(* IEC 61131-3 sources: moqui-plc/rust-plc/interfaces/plcopen-motion, 3 files *)

(* ---- types.st ---- *)
(* PLCopen Motion Control - data types used by moqui-plc.
 *
 * Interface declarations only, for type checking with a non-CODESYS compiler.
 * Names follow PLCopen Motion Control Part 1 (single axis) and Part 4
 * (coordinated motion), with the enumeration spellings used in the canonical
 * iec61131 tree. A runtime that hosts moqui-plc provides the real types.
 *
 * AXIS_REF and AXES_GROUP_REF are opaque in PLCopen; the members below are the
 * only ones the moqui-plc code reads.
 *)

TYPE AXIS_REF :
STRUCT
    wDriveId : WORD; (* drive identifier, used for log naming *)
    fTaskCycle : LREAL; (* cycle time of the motion task that runs the axis [s] *)
END_STRUCT
END_TYPE

TYPE AXES_GROUP_REF :
STRUCT
    nAxes : INT;
END_STRUCT
END_TYPE

TYPE TRIGGER_REF :
STRUCT
    iTriggerNumber : INT;
END_STRUCT
END_TYPE

TYPE MC_BUFFER_MODE : (aborting, Buffered, BlendingLow, BlendingPrevious, BlendingNext, BlendingHigh); END_TYPE
TYPE MC_DIRECTION : (negative := -1, shortest, positive, current, fastest); END_TYPE
TYPE MC_STARTMODE : (absolute, relative, ramp_in); END_TYPE
TYPE MC_TRANSITION_MODE : (TMNone, TMStartVelocity, TMConstantVelocity, TMCornerDistance, TMMaxCornerDeviation); END_TYPE
TYPE MC_CIRC_PATHCHOICE : (CLOCKWISE, COUNTER_CLOCKWISE); END_TYPE

TYPE MC_COORD_REF :
STRUCT
    X : LREAL;
    Y : LREAL;
    Z : LREAL;
    A : LREAL;
    B : LREAL;
    C : LREAL;
END_STRUCT
END_TYPE

(* Profile and cam references: content is runtime specific. *)
TYPE MC_TP_REF : STRUCT nPoints : INT; END_STRUCT END_TYPE
TYPE MC_TV_REF : STRUCT nPoints : INT; END_STRUCT END_TYPE
TYPE MC_TA_REF : STRUCT nPoints : INT; END_STRUCT END_TYPE
TYPE MC_CAM_REF : STRUCT nElements : INT; END_STRUCT END_TYPE
TYPE MC_CAM_ID : STRUCT nId : UDINT; END_STRUCT END_TYPE

(* ---- part1-single-axis.st ---- *)
(* PLCopen Motion Control Part 1 - single-axis function blocks used by moqui-plc.
 *
 * Interface declarations only (no implementation), for type checking with a
 * non-CODESYS compiler. Parameters follow the PLCopen function block
 * interface; MC_Power also carries the drive-start and regulator inputs
 * the moqui-plc code sets.
 * A runtime that hosts moqui-plc implements these blocks with the same
 * signatures.
 *)

FUNCTION_BLOCK MC_Power
VAR_IN_OUT
    Axis : AXIS_REF;
END_VAR
VAR_INPUT
    Enable : BOOL;
    bRegulatorOn : BOOL;
    bDriveStart : BOOL;
END_VAR
VAR_OUTPUT
    Status : BOOL;
    bRegulatorRealState : BOOL;
    bDriveStartRealState : BOOL;
    Busy : BOOL;
    Error : BOOL;
    ErrorID : WORD;
END_VAR
END_FUNCTION_BLOCK

FUNCTION_BLOCK MC_Home
VAR_IN_OUT
    Axis : AXIS_REF;
END_VAR
VAR_INPUT
    Execute : BOOL;
    Position : LREAL;
    BufferMode : MC_BUFFER_MODE;
END_VAR
VAR_OUTPUT
    Done : BOOL;
    Busy : BOOL;
    CommandAborted : BOOL;
    Error : BOOL;
    ErrorID : WORD;
END_VAR
END_FUNCTION_BLOCK

FUNCTION_BLOCK MC_Stop
VAR_IN_OUT
    Axis : AXIS_REF;
END_VAR
VAR_INPUT
    Execute : BOOL;
    Deceleration : LREAL;
    Jerk : LREAL;
END_VAR
VAR_OUTPUT
    Done : BOOL;
    Busy : BOOL;
    CommandAborted : BOOL;
    Error : BOOL;
    ErrorID : WORD;
END_VAR
END_FUNCTION_BLOCK

FUNCTION_BLOCK MC_Halt
VAR_IN_OUT
    Axis : AXIS_REF;
END_VAR
VAR_INPUT
    Execute : BOOL;
    Deceleration : LREAL;
    Jerk : LREAL;
    BufferMode : MC_BUFFER_MODE;
END_VAR
VAR_OUTPUT
    Done : BOOL;
    Busy : BOOL;
    Active : BOOL;
    CommandAborted : BOOL;
    Error : BOOL;
    ErrorID : WORD;
END_VAR
END_FUNCTION_BLOCK

FUNCTION_BLOCK MC_MoveAbsolute
VAR_IN_OUT
    Axis : AXIS_REF;
END_VAR
VAR_INPUT
    Execute : BOOL;
    Position : LREAL;
    Velocity : LREAL;
    Acceleration : LREAL;
    Deceleration : LREAL;
    Jerk : LREAL;
    Direction : MC_DIRECTION;
    BufferMode : MC_BUFFER_MODE;
END_VAR
VAR_OUTPUT
    Done : BOOL;
    Busy : BOOL;
    Active : BOOL;
    CommandAborted : BOOL;
    Error : BOOL;
    ErrorID : WORD;
END_VAR
END_FUNCTION_BLOCK

FUNCTION_BLOCK MC_MoveRelative
VAR_IN_OUT
    Axis : AXIS_REF;
END_VAR
VAR_INPUT
    Execute : BOOL;
    Distance : LREAL;
    Velocity : LREAL;
    Acceleration : LREAL;
    Deceleration : LREAL;
    Jerk : LREAL;
    BufferMode : MC_BUFFER_MODE;
END_VAR
VAR_OUTPUT
    Done : BOOL;
    Busy : BOOL;
    Active : BOOL;
    CommandAborted : BOOL;
    Error : BOOL;
    ErrorID : WORD;
END_VAR
END_FUNCTION_BLOCK

FUNCTION_BLOCK MC_MoveAdditive
VAR_IN_OUT
    Axis : AXIS_REF;
END_VAR
VAR_INPUT
    Execute : BOOL;
    Distance : LREAL;
    Velocity : LREAL;
    Acceleration : LREAL;
    Deceleration : LREAL;
    Jerk : LREAL;
    BufferMode : MC_BUFFER_MODE;
END_VAR
VAR_OUTPUT
    Done : BOOL;
    Busy : BOOL;
    Active : BOOL;
    CommandAborted : BOOL;
    Error : BOOL;
    ErrorID : WORD;
END_VAR
END_FUNCTION_BLOCK

FUNCTION_BLOCK MC_MoveSuperImposed
VAR_IN_OUT
    Axis : AXIS_REF;
END_VAR
VAR_INPUT
    Execute : BOOL;
    Distance : LREAL;
    VelocityDiff : LREAL;
    Acceleration : LREAL;
    Deceleration : LREAL;
    Jerk : LREAL;
END_VAR
VAR_OUTPUT
    Done : BOOL;
    Busy : BOOL;
    Active : BOOL;
    CommandAborted : BOOL;
    Error : BOOL;
    ErrorID : WORD;
END_VAR
END_FUNCTION_BLOCK

FUNCTION_BLOCK MC_HaltSuperImposed
VAR_IN_OUT
    Axis : AXIS_REF;
END_VAR
VAR_INPUT
    Execute : BOOL;
    Deceleration : LREAL;
    Jerk : LREAL;
END_VAR
VAR_OUTPUT
    Done : BOOL;
    Busy : BOOL;
    Active : BOOL;
    CommandAborted : BOOL;
    Error : BOOL;
    ErrorID : WORD;
END_VAR
END_FUNCTION_BLOCK

FUNCTION_BLOCK MC_MoveVelocity
VAR_IN_OUT
    Axis : AXIS_REF;
END_VAR
VAR_INPUT
    Execute : BOOL;
    Velocity : LREAL;
    Acceleration : LREAL;
    Deceleration : LREAL;
    Jerk : LREAL;
    Direction : MC_DIRECTION;
    BufferMode : MC_BUFFER_MODE;
END_VAR
VAR_OUTPUT
    InVelocity : BOOL;
    Busy : BOOL;
    Active : BOOL;
    CommandAborted : BOOL;
    Error : BOOL;
    ErrorID : WORD;
END_VAR
END_FUNCTION_BLOCK

FUNCTION_BLOCK MC_Jog
VAR_IN_OUT
    Axis : AXIS_REF;
END_VAR
VAR_INPUT
    JogForward : BOOL;
    JogBackward : BOOL;
    Velocity : LREAL;
    Acceleration : LREAL;
    Deceleration : LREAL;
    Jerk : LREAL;
END_VAR
VAR_OUTPUT
    Busy : BOOL;
    CommandAborted : BOOL;
    Error : BOOL;
    ErrorID : WORD;
END_VAR
END_FUNCTION_BLOCK

FUNCTION_BLOCK MC_PositionProfile
VAR_IN_OUT
    Axis : AXIS_REF;
    TimePosition : MC_TP_REF;
END_VAR
VAR_INPUT
    Execute : BOOL;
    BufferMode : MC_BUFFER_MODE;
END_VAR
VAR_OUTPUT
    Done : BOOL;
    Busy : BOOL;
    Active : BOOL;
    CommandAborted : BOOL;
    Error : BOOL;
    ErrorID : WORD;
END_VAR
END_FUNCTION_BLOCK

FUNCTION_BLOCK MC_VelocityProfile
VAR_IN_OUT
    Axis : AXIS_REF;
    TimeVelocity : MC_TV_REF;
END_VAR
VAR_INPUT
    Execute : BOOL;
    BufferMode : MC_BUFFER_MODE;
END_VAR
VAR_OUTPUT
    Done : BOOL;
    Busy : BOOL;
    Active : BOOL;
    CommandAborted : BOOL;
    Error : BOOL;
    ErrorID : WORD;
END_VAR
END_FUNCTION_BLOCK

FUNCTION_BLOCK MC_AccelerationProfile
VAR_IN_OUT
    Axis : AXIS_REF;
    TimeAcceleration : MC_TA_REF;
END_VAR
VAR_INPUT
    Execute : BOOL;
    BufferMode : MC_BUFFER_MODE;
END_VAR
VAR_OUTPUT
    Done : BOOL;
    Busy : BOOL;
    Active : BOOL;
    CommandAborted : BOOL;
    Error : BOOL;
    ErrorID : WORD;
END_VAR
END_FUNCTION_BLOCK

FUNCTION_BLOCK MC_SetPosition
VAR_IN_OUT
    Axis : AXIS_REF;
END_VAR
VAR_INPUT
    Execute : BOOL;
    Position : LREAL;
    Mode : BOOL;
END_VAR
VAR_OUTPUT
    Done : BOOL;
    Busy : BOOL;
    Error : BOOL;
    ErrorID : WORD;
END_VAR
END_FUNCTION_BLOCK

FUNCTION_BLOCK MC_SetOverride
VAR_IN_OUT
    Axis : AXIS_REF;
END_VAR
VAR_INPUT
    Enable : BOOL;
    VelFactor : LREAL;
    AccFactor : LREAL;
    JerkFactor : LREAL;
END_VAR
VAR_OUTPUT
    Enabled : BOOL;
    Busy : BOOL;
    Error : BOOL;
    ErrorID : WORD;
END_VAR
END_FUNCTION_BLOCK

FUNCTION_BLOCK MC_ReadParameter
VAR_IN_OUT
    Axis : AXIS_REF;
END_VAR
VAR_INPUT
    Enable : BOOL;
    ParameterNumber : DINT;
END_VAR
VAR_OUTPUT
    Valid : BOOL;
    Busy : BOOL;
    Error : BOOL;
    ErrorID : WORD;
    Value : LREAL;
END_VAR
END_FUNCTION_BLOCK

FUNCTION_BLOCK MC_ReadBoolParameter
VAR_IN_OUT
    Axis : AXIS_REF;
END_VAR
VAR_INPUT
    Enable : BOOL;
    ParameterNumber : DINT;
END_VAR
VAR_OUTPUT
    Valid : BOOL;
    Busy : BOOL;
    Error : BOOL;
    ErrorID : WORD;
    Value : BOOL;
END_VAR
END_FUNCTION_BLOCK

FUNCTION_BLOCK MC_WriteParameter
VAR_IN_OUT
    Axis : AXIS_REF;
END_VAR
VAR_INPUT
    Execute : BOOL;
    ParameterNumber : DINT;
    Value : LREAL;
END_VAR
VAR_OUTPUT
    Done : BOOL;
    Busy : BOOL;
    Error : BOOL;
    ErrorID : WORD;
END_VAR
END_FUNCTION_BLOCK

FUNCTION_BLOCK MC_WriteBoolParameter
VAR_IN_OUT
    Axis : AXIS_REF;
END_VAR
VAR_INPUT
    Execute : BOOL;
    ParameterNumber : DINT;
    Value : BOOL;
END_VAR
VAR_OUTPUT
    Done : BOOL;
    Busy : BOOL;
    Error : BOOL;
    ErrorID : WORD;
END_VAR
END_FUNCTION_BLOCK

FUNCTION_BLOCK MC_ReadActualPosition
VAR_IN_OUT
    Axis : AXIS_REF;
END_VAR
VAR_INPUT
    Enable : BOOL;
END_VAR
VAR_OUTPUT
    Valid : BOOL;
    Busy : BOOL;
    Error : BOOL;
    ErrorID : WORD;
    Position : LREAL;
END_VAR
END_FUNCTION_BLOCK

FUNCTION_BLOCK MC_ReadActualVelocity
VAR_IN_OUT
    Axis : AXIS_REF;
END_VAR
VAR_INPUT
    Enable : BOOL;
END_VAR
VAR_OUTPUT
    Valid : BOOL;
    Busy : BOOL;
    Error : BOOL;
    ErrorID : WORD;
    Velocity : LREAL;
END_VAR
END_FUNCTION_BLOCK

FUNCTION_BLOCK MC_ReadActualTorque
VAR_IN_OUT
    Axis : AXIS_REF;
END_VAR
VAR_INPUT
    Enable : BOOL;
END_VAR
VAR_OUTPUT
    Valid : BOOL;
    Busy : BOOL;
    Error : BOOL;
    ErrorID : WORD;
    Torque : LREAL;
END_VAR
END_FUNCTION_BLOCK

FUNCTION_BLOCK MC_ReadStatus
VAR_IN_OUT
    Axis : AXIS_REF;
END_VAR
VAR_INPUT
    Enable : BOOL;
END_VAR
VAR_OUTPUT
    Valid : BOOL;
    Busy : BOOL;
    Error : BOOL;
    ErrorID : WORD;
    ErrorStop : BOOL;
    Disabled : BOOL;
    Stopping : BOOL;
    Homing : BOOL;
    Standstill : BOOL;
    DiscreteMotion : BOOL;
    ContinuousMotion : BOOL;
    SynchronizedMotion : BOOL;
END_VAR
END_FUNCTION_BLOCK

FUNCTION_BLOCK MC_ReadAxisError
VAR_IN_OUT
    Axis : AXIS_REF;
END_VAR
VAR_INPUT
    Enable : BOOL;
END_VAR
VAR_OUTPUT
    Valid : BOOL;
    Busy : BOOL;
    Error : BOOL;
    ErrorID : WORD;
    AxisErrorID : DWORD;
END_VAR
END_FUNCTION_BLOCK

FUNCTION_BLOCK MC_Reset
VAR_IN_OUT
    Axis : AXIS_REF;
END_VAR
VAR_INPUT
    Execute : BOOL;
END_VAR
VAR_OUTPUT
    Done : BOOL;
    Busy : BOOL;
    Error : BOOL;
    ErrorID : WORD;
END_VAR
END_FUNCTION_BLOCK

FUNCTION_BLOCK MC_TouchProbe
VAR_IN_OUT
    Axis : AXIS_REF;
    TriggerInput : TRIGGER_REF;
END_VAR
VAR_INPUT
    Execute : BOOL;
    WindowOnly : BOOL;
    FirstPosition : LREAL;
    LastPosition : LREAL;
END_VAR
VAR_OUTPUT
    Done : BOOL;
    Busy : BOOL;
    CommandAborted : BOOL;
    Error : BOOL;
    ErrorID : WORD;
    RecordedPosition : LREAL;
END_VAR
END_FUNCTION_BLOCK

FUNCTION_BLOCK MC_AbortTrigger
VAR_IN_OUT
    Axis : AXIS_REF;
    TriggerInput : TRIGGER_REF;
END_VAR
VAR_INPUT
    Execute : BOOL;
END_VAR
VAR_OUTPUT
    Done : BOOL;
    Busy : BOOL;
    Error : BOOL;
    ErrorID : WORD;
END_VAR
END_FUNCTION_BLOCK

FUNCTION_BLOCK MC_CamTableSelect
VAR_IN_OUT
    Master : AXIS_REF;
    Slave : AXIS_REF;
    CamTable : MC_CAM_REF;
END_VAR
VAR_INPUT
    Execute : BOOL;
    Periodic : BOOL;
    MasterAbsolute : BOOL;
    SlaveAbsolute : BOOL;
END_VAR
VAR_OUTPUT
    Done : BOOL;
    Busy : BOOL;
    Error : BOOL;
    ErrorID : WORD;
    CamTableID : MC_CAM_ID;
END_VAR
END_FUNCTION_BLOCK

FUNCTION_BLOCK MC_CamIn
VAR_IN_OUT
    Master : AXIS_REF;
    Slave : AXIS_REF;
END_VAR
VAR_INPUT
    Execute : BOOL;
    MasterOffset : LREAL;
    SlaveOffset : LREAL;
    MasterScaling : LREAL;
    SlaveScaling : LREAL;
    StartMode : MC_STARTMODE;
    CamTableID : MC_CAM_ID;
    BufferMode : MC_BUFFER_MODE;
END_VAR
VAR_OUTPUT
    InSync : BOOL;
    Busy : BOOL;
    Active : BOOL;
    CommandAborted : BOOL;
    Error : BOOL;
    ErrorID : WORD;
    EndOfProfile : BOOL;
END_VAR
END_FUNCTION_BLOCK

FUNCTION_BLOCK MC_CamOut
VAR_IN_OUT
    Slave : AXIS_REF;
END_VAR
VAR_INPUT
    Execute : BOOL;
END_VAR
VAR_OUTPUT
    Done : BOOL;
    Busy : BOOL;
    Error : BOOL;
    ErrorID : WORD;
END_VAR
END_FUNCTION_BLOCK

FUNCTION_BLOCK MC_GearIn
VAR_IN_OUT
    Master : AXIS_REF;
    Slave : AXIS_REF;
END_VAR
VAR_INPUT
    Execute : BOOL;
    RatioNumerator : DINT;
    RatioDenominator : UDINT;
    Acceleration : LREAL;
    Deceleration : LREAL;
    Jerk : LREAL;
    BufferMode : MC_BUFFER_MODE;
END_VAR
VAR_OUTPUT
    InGear : BOOL;
    Busy : BOOL;
    Active : BOOL;
    CommandAborted : BOOL;
    Error : BOOL;
    ErrorID : WORD;
END_VAR
END_FUNCTION_BLOCK

FUNCTION_BLOCK MC_GearInPos
VAR_IN_OUT
    Master : AXIS_REF;
    Slave : AXIS_REF;
END_VAR
VAR_INPUT
    Execute : BOOL;
    RatioNumerator : DINT;
    RatioDenominator : UDINT;
    MasterSyncPosition : LREAL;
    SlaveSyncPosition : LREAL;
    MasterStartDistance : LREAL;
    Velocity : LREAL;
    Acceleration : LREAL;
    Deceleration : LREAL;
    Jerk : LREAL;
    BufferMode : MC_BUFFER_MODE;
END_VAR
VAR_OUTPUT
    StartSync : BOOL;
    InSync : BOOL;
    Busy : BOOL;
    Active : BOOL;
    CommandAborted : BOOL;
    Error : BOOL;
    ErrorID : WORD;
END_VAR
END_FUNCTION_BLOCK

FUNCTION_BLOCK MC_GearOut
VAR_IN_OUT
    Slave : AXIS_REF;
END_VAR
VAR_INPUT
    Execute : BOOL;
END_VAR
VAR_OUTPUT
    Done : BOOL;
    Busy : BOOL;
    Error : BOOL;
    ErrorID : WORD;
END_VAR
END_FUNCTION_BLOCK

FUNCTION_BLOCK MC_Phasing
VAR_IN_OUT
    Master : AXIS_REF;
    Slave : AXIS_REF;
END_VAR
VAR_INPUT
    Execute : BOOL;
    PhaseShift : LREAL;
    Velocity : LREAL;
    Acceleration : LREAL;
    Deceleration : LREAL;
    Jerk : LREAL;
    BufferMode : MC_BUFFER_MODE;
END_VAR
VAR_OUTPUT
    Done : BOOL;
    Busy : BOOL;
    Active : BOOL;
    CommandAborted : BOOL;
    Error : BOOL;
    ErrorID : WORD;
END_VAR
END_FUNCTION_BLOCK

(* ---- part4-coordinated.st ---- *)
(* PLCopen Motion Control Part 4 - axis group function blocks used by moqui-plc.
 *
 * Interface declarations only (no implementation), for type checking with a
 * non-CODESYS compiler. Parameters follow the PLCopen function block
 * interface; positions use SMC_POS_REF, the CODESYS position type
 * (codesys-softmotion/softmotion.st).
 * A runtime that hosts moqui-plc implements these blocks with the same
 * signatures.
 *)

FUNCTION_BLOCK MC_GroupEnable
VAR_IN_OUT
    AxisGroup : AXES_GROUP_REF;
END_VAR
VAR_INPUT
    Execute : BOOL;
END_VAR
VAR_OUTPUT
    Done : BOOL;
    Busy : BOOL;
    Error : BOOL;
    ErrorID : WORD;
END_VAR
END_FUNCTION_BLOCK

FUNCTION_BLOCK MC_GroupReset
VAR_IN_OUT
    AxisGroup : AXES_GROUP_REF;
END_VAR
VAR_INPUT
    Execute : BOOL;
END_VAR
VAR_OUTPUT
    Done : BOOL;
    Busy : BOOL;
    Error : BOOL;
    ErrorID : WORD;
END_VAR
END_FUNCTION_BLOCK

FUNCTION_BLOCK MC_GroupStop
VAR_IN_OUT
    AxisGroup : AXES_GROUP_REF;
END_VAR
VAR_INPUT
    Execute : BOOL;
    Deceleration : LREAL;
    Jerk : LREAL;
END_VAR
VAR_OUTPUT
    Done : BOOL;
    Busy : BOOL;
    CommandAborted : BOOL;
    Error : BOOL;
    ErrorID : WORD;
END_VAR
END_FUNCTION_BLOCK

FUNCTION_BLOCK MC_GroupHalt
VAR_IN_OUT
    AxisGroup : AXES_GROUP_REF;
END_VAR
VAR_INPUT
    Execute : BOOL;
    Deceleration : LREAL;
    Jerk : LREAL;
    AccFactor : LREAL;
    JerkFactor : LREAL;
    BufferMode : MC_BUFFER_MODE;
END_VAR
VAR_OUTPUT
    Done : BOOL;
    Busy : BOOL;
    Active : BOOL;
    CommandAborted : BOOL;
    Error : BOOL;
    ErrorID : WORD;
END_VAR
END_FUNCTION_BLOCK

FUNCTION_BLOCK MC_GroupSetOverride
VAR_IN_OUT
    AxisGroup : AXES_GROUP_REF;
END_VAR
VAR_INPUT
    Enable : BOOL;
    VelFactor : LREAL;
    AccFactor : LREAL;
    JerkFactor : LREAL;
END_VAR
VAR_OUTPUT
    Enabled : BOOL;
    Busy : BOOL;
    Error : BOOL;
    ErrorID : WORD;
END_VAR
END_FUNCTION_BLOCK

FUNCTION_BLOCK MC_GroupReadActualPosition
VAR_IN_OUT
    AxisGroup : AXES_GROUP_REF;
END_VAR
VAR_INPUT
    Enable : BOOL;
    CoordSystem : SMC_COORD_SYSTEM;
END_VAR
VAR_OUTPUT
    Valid : BOOL;
    Busy : BOOL;
    Error : BOOL;
    ErrorID : WORD;
    Position : SMC_POS_REF;
END_VAR
END_FUNCTION_BLOCK

FUNCTION_BLOCK MC_GroupReadActualVelocity
VAR_IN_OUT
    AxisGroup : AXES_GROUP_REF;
END_VAR
VAR_INPUT
    Enable : BOOL;
    CoordSystem : SMC_COORD_SYSTEM;
END_VAR
VAR_OUTPUT
    Valid : BOOL;
    Busy : BOOL;
    Error : BOOL;
    ErrorID : WORD;
    Velocity : SMC_POS_REF;
END_VAR
END_FUNCTION_BLOCK

FUNCTION_BLOCK MC_GroupReadError
VAR_IN_OUT
    AxisGroup : AXES_GROUP_REF;
END_VAR
VAR_INPUT
    Enable : BOOL;
END_VAR
VAR_OUTPUT
    Valid : BOOL;
    Busy : BOOL;
    Error : BOOL;
    ErrorID : WORD;
    GroupErrorID : DWORD;
END_VAR
END_FUNCTION_BLOCK

FUNCTION_BLOCK MC_GroupReadStatus
VAR_IN_OUT
    AxisGroup : AXES_GROUP_REF;
END_VAR
VAR_INPUT
    Enable : BOOL;
END_VAR
VAR_OUTPUT
    Valid : BOOL;
    Busy : BOOL;
    Error : BOOL;
    ErrorID : WORD;
    GroupMoving : BOOL;
    GroupHoming : BOOL;
    GroupErrorStop : BOOL;
    GroupStandby : BOOL;
    GroupStopping : BOOL;
    GroupDisabled : BOOL;
END_VAR
END_FUNCTION_BLOCK

FUNCTION_BLOCK MC_MoveLinearAbsolute
VAR_IN_OUT
    AxisGroup : AXES_GROUP_REF;
END_VAR
VAR_INPUT
    Execute : BOOL;
    Position : SMC_POS_REF;
    Velocity : LREAL;
    Acceleration : LREAL;
    Deceleration : LREAL;
    Jerk : LREAL;
    CoordSystem : SMC_COORD_SYSTEM;
    BufferMode : MC_BUFFER_MODE;
    TransitionMode : MC_TRANSITION_MODE;
    TransitionParameter : ARRAY [0..(SMC_RCNST.MAX_TRANS_PARAMS - 1)] OF LREAL;
END_VAR
VAR_OUTPUT
    Done : BOOL;
    Busy : BOOL;
    Active : BOOL;
    CommandAborted : BOOL;
    Error : BOOL;
    ErrorID : WORD;
END_VAR
END_FUNCTION_BLOCK

FUNCTION_BLOCK MC_MoveLinearRelative
VAR_IN_OUT
    AxisGroup : AXES_GROUP_REF;
END_VAR
VAR_INPUT
    Execute : BOOL;
    Distance : SMC_POS_REF;
    Velocity : LREAL;
    Acceleration : LREAL;
    Deceleration : LREAL;
    Jerk : LREAL;
    CoordSystem : SMC_COORD_SYSTEM;
    BufferMode : MC_BUFFER_MODE;
    TransitionMode : MC_TRANSITION_MODE;
    TransitionParameter : ARRAY [0..(SMC_RCNST.MAX_TRANS_PARAMS - 1)] OF LREAL;
END_VAR
VAR_OUTPUT
    Done : BOOL;
    Busy : BOOL;
    Active : BOOL;
    CommandAborted : BOOL;
    Error : BOOL;
    ErrorID : WORD;
END_VAR
END_FUNCTION_BLOCK

FUNCTION_BLOCK MC_MoveDirectAbsolute
VAR_IN_OUT
    AxisGroup : AXES_GROUP_REF;
END_VAR
VAR_INPUT
    Execute : BOOL;
    Position : SMC_POS_REF;
    CoordSystem : SMC_COORD_SYSTEM;
    BufferMode : MC_BUFFER_MODE;
    TransitionMode : MC_TRANSITION_MODE;
    TransitionParameter : ARRAY [0..(SMC_RCNST.MAX_TRANS_PARAMS - 1)] OF LREAL;
END_VAR
VAR_OUTPUT
    Done : BOOL;
    Busy : BOOL;
    Active : BOOL;
    CommandAborted : BOOL;
    Error : BOOL;
    ErrorID : WORD;
END_VAR
END_FUNCTION_BLOCK

FUNCTION_BLOCK MC_MoveDirectRelative
VAR_IN_OUT
    AxisGroup : AXES_GROUP_REF;
END_VAR
VAR_INPUT
    Execute : BOOL;
    Distance : SMC_POS_REF;
    CoordSystem : SMC_COORD_SYSTEM;
    BufferMode : MC_BUFFER_MODE;
    TransitionMode : MC_TRANSITION_MODE;
    TransitionParameter : ARRAY [0..(SMC_RCNST.MAX_TRANS_PARAMS - 1)] OF LREAL;
END_VAR
VAR_OUTPUT
    Done : BOOL;
    Busy : BOOL;
    Active : BOOL;
    CommandAborted : BOOL;
    Error : BOOL;
    ErrorID : WORD;
END_VAR
END_FUNCTION_BLOCK

FUNCTION_BLOCK MC_MoveCircularAbsolute
VAR_IN_OUT
    AxisGroup : AXES_GROUP_REF;
END_VAR
VAR_INPUT
    Execute : BOOL;
    CircMode : SMC_CIRC_MODE;
    AuxPoint : SMC_POS_REF;
    EndPoint : SMC_POS_REF;
    PathChoice : MC_CIRC_PATHCHOICE;
    Velocity : LREAL;
    Acceleration : LREAL;
    Deceleration : LREAL;
    Jerk : LREAL;
    CoordSystem : SMC_COORD_SYSTEM;
    BufferMode : MC_BUFFER_MODE;
    TransitionMode : MC_TRANSITION_MODE;
    TransitionParameter : ARRAY [0..(SMC_RCNST.MAX_TRANS_PARAMS - 1)] OF LREAL;
END_VAR
VAR_OUTPUT
    Done : BOOL;
    Busy : BOOL;
    Active : BOOL;
    CommandAborted : BOOL;
    Error : BOOL;
    ErrorID : WORD;
END_VAR
END_FUNCTION_BLOCK

FUNCTION_BLOCK MC_MoveCircularRelative
VAR_IN_OUT
    AxisGroup : AXES_GROUP_REF;
END_VAR
VAR_INPUT
    Execute : BOOL;
    CircMode : SMC_CIRC_MODE;
    AuxPoint : SMC_POS_REF;
    EndPoint : SMC_POS_REF;
    PathChoice : MC_CIRC_PATHCHOICE;
    Velocity : LREAL;
    Acceleration : LREAL;
    Deceleration : LREAL;
    Jerk : LREAL;
    CoordSystem : SMC_COORD_SYSTEM;
    BufferMode : MC_BUFFER_MODE;
    TransitionMode : MC_TRANSITION_MODE;
    TransitionParameter : ARRAY [0..(SMC_RCNST.MAX_TRANS_PARAMS - 1)] OF LREAL;
END_VAR
VAR_OUTPUT
    Done : BOOL;
    Busy : BOOL;
    Active : BOOL;
    CommandAborted : BOOL;
    Error : BOOL;
    ErrorID : WORD;
END_VAR
END_FUNCTION_BLOCK

FUNCTION_BLOCK MC_SetCoordinateTransform
VAR_IN_OUT
    AxisGroup : AXES_GROUP_REF;
END_VAR
VAR_INPUT
    Execute : BOOL;
    CoordSystem : SMC_COORD_SYSTEM;
    CoordTransform : MC_COORD_REF;
    BufferMode : MC_BUFFER_MODE;
END_VAR
VAR_OUTPUT
    Done : BOOL;
    Busy : BOOL;
    Error : BOOL;
    ErrorID : WORD;
END_VAR
END_FUNCTION_BLOCK

FUNCTION_BLOCK MC_TrackConveyorBelt
VAR_IN_OUT
    AxisGroup : AXES_GROUP_REF;
    ConveyorBelt : AXIS_REF;
END_VAR
VAR_INPUT
    Execute : BOOL;
    ConveyorBeltOrigin : MC_COORD_REF;
    InitialObjectPosition : MC_COORD_REF;
    CoordSystem : SMC_COORD_SYSTEM;
END_VAR
VAR_OUTPUT
    Done : BOOL;
    Busy : BOOL;
    Error : BOOL;
    ErrorID : WORD;
    cs : SMC_CoordinateSystem;
END_VAR
END_FUNCTION_BLOCK

FUNCTION_BLOCK MC_TrackRotaryTable
VAR_IN_OUT
    AxisGroup : AXES_GROUP_REF;
    RotaryTable : AXIS_REF;
END_VAR
VAR_INPUT
    Execute : BOOL;
    RotaryTableOrigin : MC_COORD_REF;
    InitialObjectPosition : MC_COORD_REF;
    CoordSystem : SMC_COORD_SYSTEM;
END_VAR
VAR_OUTPUT
    Done : BOOL;
    Busy : BOOL;
    Error : BOOL;
    ErrorID : WORD;
    cs : SMC_CoordinateSystem;
END_VAR
END_FUNCTION_BLOCK
